FUNCTION_BLOCK PID_LOOP (* Migrated from IEC 61131-3 ST *)
  (* Standard: 61499-2 *)
  (* Version 1.0, 2026-11-06, st2fb *)
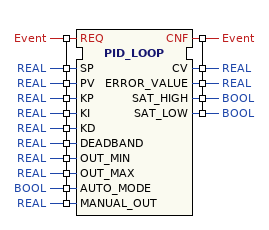
  EVENT_INPUT
    REQ WITH SP, PV, KP, KI, KD, DEADBAND, OUT_MIN, OUT_MAX, AUTO_MODE, MANUAL_OUT;
  END_EVENT
  EVENT_OUTPUT
    CNF WITH CV, ERROR_VALUE, SAT_HIGH, SAT_LOW;
  END_EVENT
  VAR_INPUT
    SP : REAL;
    PV : REAL;
    KP : REAL;
    KI : REAL;
    KD : REAL;
    DEADBAND : REAL;
    OUT_MIN : REAL;
    OUT_MAX : REAL;
    AUTO_MODE : BOOL;
    MANUAL_OUT : REAL;
  END_VAR
  VAR_OUTPUT
    CV : REAL;
    ERROR_VALUE : REAL;
    SAT_HIGH : BOOL;
    SAT_LOW : BOOL;
  END_VAR
  VAR
    I_TERM : REAL;
    PREV_PV : REAL;
    UNCLAMPED : REAL;
  END_VAR
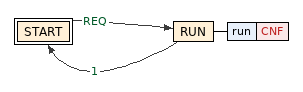
  EC_STATES
    START;
    RUN : run -> CNF;
  END_STATES
  EC_TRANSITIONS
    START TO RUN := REQ;
    RUN TO START := 1;
  END_TRANSITIONS
  ALGORITHM run IN ST:
ERROR_VALUE := SP - PV;
IF (ERROR_VALUE < DEADBAND) AND (ERROR_VALUE > 0.0 - DEADBAND) THEN
  ERROR_VALUE := 0.0;
END_IF;
IF AUTO_MODE THEN
  IF NOT ((SAT_HIGH AND ERROR_VALUE > 0.0) OR (SAT_LOW AND ERROR_VALUE < 0.0)) THEN
    I_TERM := I_TERM + KI * ERROR_VALUE;
  END_IF;
  UNCLAMPED := KP * ERROR_VALUE + I_TERM - KD * (PV - PREV_PV);
ELSE
  UNCLAMPED := MANUAL_OUT;
  I_TERM := MANUAL_OUT - KP * ERROR_VALUE;
END_IF;
SAT_HIGH := UNCLAMPED >= OUT_MAX;
SAT_LOW := UNCLAMPED <= OUT_MIN;
IF SAT_HIGH THEN
  CV := OUT_MAX;
ELSIF SAT_LOW THEN
  CV := OUT_MIN;
ELSE
  CV := UNCLAMPED;
END_IF;
PREV_PV := PV;
  END_ALGORITHM
END_FUNCTION_BLOCK
